FUNCTION_BLOCK FB_CoverIdleState EXTENDS FB_CoverState
VAR_INPUT
END_VAR
VAR_OUTPUT
END_VAR
VAR
END_VAR

METHOD CloseCommand : BOOL
pCover^.SetState(pCover^.fbCoverClosingState);
END_METHOD

METHOD OpenCommand : BOOL
pCover^.SetState(pCover^.fbCoverOpeningState);
END_METHOD

METHOD StopCommand : BOOL
pCover^.SetState(pCover^.fbCoverStoppingState);
END_METHOD

END_FUNCTION_BLOCK

(* stored: Version 1.1.0.1, ProductVersion 3.1.4024.15
   POU FB_CoverIdleState: Id {f1d58d15-5a8c-4164-99e1-a5d9e089ed6c}, SpecialFunc None
   Method CloseCommand: Id {6dfe491a-a1e5-4076-a615-62fc471ebe72}
   Method OpenCommand: Id {4c8f3564-fa75-48d7-b56e-701d8b57a66d}
   Method StopCommand: Id {43efa24f-8021-4279-87de-321de14fc42b} *)
